(* IEC 61131-3 sources: genai_codesys/experiments/raw/formal/20261109_234635_2ba96d/public_02/codex_cli__deepseek-v4.1-flash-1017/attempt_00, 2 files *)

(* ---- declaration.st ---- *)
FUNCTION_BLOCK FB_DWordEdgeDetection
VAR_INPUT
    value : DWORD;
END_VAR
VAR_OUTPUT
    hasChanged : BOOL;
    hasRisingEdges : BOOL;
    risingBits : DWORD;
    noOfRisingBits : USINT;
    hasFallingEdges : BOOL;
    fallingBits : DWORD;
    noOfFallingBits : USINT;
END_VAR
VAR
    lastValue : DWORD;
    i : INT;
END_VAR
END_FUNCTION_BLOCK

(* ---- implementation.st ---- *)
hasChanged := value <> lastValue;

risingBits := value AND NOT lastValue;
fallingBits := lastValue AND NOT value;

hasRisingEdges := risingBits <> DWORD#0;
hasFallingEdges := fallingBits <> DWORD#0;

noOfRisingBits := 0;
noOfFallingBits := 0;

FOR i := 0 TO 31 DO
    IF (risingBits AND SHL(DWORD#1, i)) <> DWORD#0 THEN
        noOfRisingBits := noOfRisingBits + 1;
    END_IF;

    IF (fallingBits AND SHL(DWORD#1, i)) <> DWORD#0 THEN
        noOfFallingBits := noOfFallingBits + 1;
    END_IF;
END_FOR;

lastValue := value;
